// TIA Portal V21 export
// export: Created 2026-11-21T13:31:41.3940929Z, ExportSetting WithDefaults, DisplayName Totally Integrated Automation Portal, DisplayVersion V21, DisplayName STEP 7 Professional, DisplayVersion V21, DisplayName STEP 7 Safety, DisplayVersion V21, DisplayName Tech WebApplication, DisplayVersion V21, DisplayName WinCC Basic/Comfort/Advanced, DisplayVersion V21, DisplayName WinCC Unified, DisplayVersion V21
VAR_GLOBAL   // PLC tag table "Default tag table"
   Tag__639308646888752274 AT %T1 : Timer;
   Tag__639308646889222918 AT %I0.2 : Bool;
   Tag__639308646889222919 AT %C1 : Counter;
   Tag__639308646889222920 AT %I0.3 : Bool;
   Tag__639308646889546626 AT %MW10 : Word;
   Tag__639308646889705153 AT %QW0 : Word;
END_VAR
